PROGRAM MAIN
VAR
	
tempVar			: BOOL;

END_VAR

END_PROGRAM

(* stored: Version 1.1.0.1
   POU MAIN: Id {29a5c702-63ab-46b2-8e24-c0f72590d031}, SpecialFunc None *)
